// TIA Portal V20 export
// export: Created 2026-10-12T16:46:22.8168119Z, ExportSetting WithDefaults, DisplayName Totally Integrated Automation Portal, DisplayVersion V20 Update 6, DisplayName TIA Portal Openness, DisplayVersion V20 Update 6, DisplayName TIA Portal Version Control Interface, DisplayVersion V20 Update 6, DisplayName SINAMICS Startdrive Advanced, DisplayVersion V20 SP1 Update 2, DisplayName SINAMICS Startdrive G110M, G120, G120C, G120D, G120P, G115D, DisplayVersion V20 SP1 Update 2, DisplayName SINAMICS Startdrive G130, G150, S120, S150, SINAMICS MV, G220, S200, S210, DisplayVersion V20 SP1 Update 2, DisplayName STEP 7 Professional, DisplayVersion V20 Update 6, DisplayName STEP 7 Safety, DisplayVersion V20 Update 2, DisplayName WinCC Basic/Comfort/Advanced, DisplayVersion V20 Update 6, DisplayName WinCC Professional, DisplayVersion V20 Update 6, DisplayName WinCC Unified, DisplayVersion V20 Update 6
TYPE "UDT_Bad_Konfig"
// stored: IsFailsafeCompliant false
   STRUCT
      Ausstattung : Struct
         HatHeizung_1 { S7_SetPoint := 'True'} : Bool;
         HatHeizung_2 { S7_SetPoint := 'True'} : Bool;
         HatPumpe { S7_SetPoint := 'True'} : Bool;
         HatPumpe_FU { S7_SetPoint := 'True'} : Bool;
         HatWarenbewegung_X { S7_SetPoint := 'True'} : Bool;
         HatWarenbewegung_Y { S7_SetPoint := 'True'} : Bool;
         HatUltraschall { S7_SetPoint := 'True'} : Bool;
         HatGleichrichter { S7_SetPoint := 'True'} : Bool;
         HatNiveau { S7_SetPoint := 'True'} : Bool;
      END_STRUCT;
      IO_Ein : Struct
         WT_Einsetzen : Array[1..3] of Bool;
         WT_Entnehmen : Array[1..3] of Bool;
         Ist_Temperatur_1 : Real;
         Ist_Temperatur_2 : Real;
         Niveau_OK : Bool;
         Motorschutz_OK : Bool;
         FI_Schutz_OK : Bool;
         Kein_Uebertemp : Bool;
         FU_Pumpe_Bereit : Bool;
         FU_WB1_Bereit : Bool;
         FU_WB2_Bereit : Bool;
      END_STRUCT;
      IO_Aus : Struct
         Ampel_Gruen : Bool;
         Ampel_Orange : Bool;
         Ampel_Rot : Bool;
         Pumpe : Bool;
         Pumpe_FU_Freigabe : Bool;
         Pumpe_FU_Netzschuetz : Bool;
         Pumpe_FU_Reset : Bool;
         Heizung_1_Regelung : Bool;
         Heizung_1_Sicherheit : Bool;
         Heizung_2_Regelung : Bool;
         Heizung_2_Sicherheit : Bool;
         Ultraschall_Freigabe : Bool;
         LED_Einsetzen : Array[1..3] of Bool;
         LED_Entnehmen : Array[1..3] of Bool;
         LED_Vorwarn : Array[1..3] of Bool;
         LED_Heizung_Aktiv : Bool;
         LED_Stoerung : Bool;
         LED_Handbetrieb : Bool;
         Prio_Einsetzen_WT : Int;
         Prio_Entnehmen_WT : Int;
      END_STRUCT;
      Pumpe_Ein : Bool;
      Pumpe_FU_Soll : Real;
      Ultraschall_Ein : Bool;
      Heizung_1_Soll : Real;
      Heizung_1_Ist : Real;
      Heizung_2_Soll : Real;
      Heizung_2_Ist : Real;
      Warenbewegung_X_Soll : Real;
      Warenbewegung_X_Ist : Real;
      Warenbewegung_Y_Soll : Real;
      Warenbewegung_Y_Ist : Real;
      WB1_Reset : Bool;
      WB2_Reset : Bool;
      GR_Aktiv : Bool;
      GR_Strom_Soll : Real;
      GR_Strom_Ist : Real;
      GR_Spannung_Soll : Real;
      GR_Spannung_Ist : Real;
      GR_Pulsfrequenz : Real;
      GR_DutyCycle : Real;
      WT { S7_SetPoint := 'True'} : Array[1..3] of "UDT_WT_Platz";
      Ampel_Status : Int;
      Hupe : Bool;
      Betriebsbereit : Bool;
      Hand_Aktiv_Intern : Bool;
      FU_Pumpe_Stoerung : Bool;
      FU_WB1_Stoerung : Bool;
      FU_WB2_Stoerung : Bool;
   END_STRUCT;
END_TYPE
